// TIA Portal V21 export
// export: Created 2026-08-21T20:18:56.7269124Z, ExportSetting None, DisplayName Totally Integrated Automation Portal, DisplayVersion V21, DisplayName STEP 7 Professional, DisplayVersion V21, DisplayName STEP 7 Safety, DisplayVersion V21, DisplayName Tech WebApplication, DisplayVersion V21, DisplayName WinCC Basic/Comfort/Advanced, DisplayVersion V21, DisplayName WinCC Professional, DisplayVersion V21, DisplayName WinCC Unified, DisplayVersion V21
TYPE "UDT_Service_StepMedium"
   STRUCT
      command : Array[0..0] of DWord;   // 'Command' configuration of control modules for sequencer
      force : Array[0..0] of DWord;   // 'Force' configuration of control modules for sequencer
      check : Array[0..0] of DWord;   // 'Check' configuration of control modules for sequencer
      "or" : Array[0..0] of DWord;   // Logical 'OR' configuration of control modules for sequencer
   END_STRUCT;
   // command[0] := 16#FFFFFFFF;
   // force[0] := 16#FFFFFFFF;
   // check[0] := 16#FFFFFFFF;
   // "or"[0] := 16#FFFFFFFF;
END_TYPE
